TYPE ST_SFC :
STRUCT
	SFCInit:		REFERENCE TO BOOL;
	SFCReset:		REFERENCE TO BOOL;
	SFCError:		REFERENCE TO BOOL;
	SFCEnableLimit:	REFERENCE TO BOOL;
	SFCErrorStep:	REFERENCE TO STRING;
	SFCErrorPOU:	REFERENCE TO STRING;
	SFCQuitError:	REFERENCE TO BOOL;
	SFCPause:		REFERENCE TO BOOL;
	SFCTrans:		REFERENCE TO BOOL;
	SFCCurrentStep:	REFERENCE TO STRING;
	SFCTip:			REFERENCE TO BOOL;
	SFCTipMode:		REFERENCE TO BOOL;
END_STRUCT
END_TYPE

(* stored: Version 1.1.0.1, ProductVersion 3.1.4024.12
   DUT ST_SFC: Id {f04d6c9c-5a02-439c-baf9-fe585b1e25a6} *)
